(* IEC 61131-3 sources: STAR-PLC-Agent/experiments/E3/campaign_2026-11-14T074447614126+0000/PUB003/run_2026-11-14T075406993896+0000/compile_00, 1 file *)

(* ---- FB_Task.st ---- *)
FUNCTION_BLOCK FB_Task
VAR_INPUT
    Value : REAL;
    hiLevel : REAL;
    loLevel : REAL;
    hystWindow : REAL;
END_VAR
VAR_OUTPUT
    hiAlarm : BOOL := FALSE;
    loAlarm : BOOL := FALSE;
    {attribute 'analysis' := '-27'}
    error : BOOL := FALSE;
    {attribute 'analysis' := '-27'}
    status : WORD := 0;
END_VAR
VAR
    hiAlarmState : BOOL := FALSE;
    loAlarmState : BOOL := FALSE;
    span : REAL;
    hiRelease : REAL;
    loRelease : REAL;
END_VAR

span := hiLevel - loLevel;
hiRelease := hiLevel - hystWindow;
loRelease := loLevel + hystWindow;

IF loLevel >= hiLevel THEN
    error := TRUE;
    status := 16#8001;
ELSIF hystWindow >= span THEN
    error := TRUE;
    status := 16#8002;
ELSE
    error := FALSE;
    status := 0;

    IF Value > hiLevel THEN
        hiAlarmState := TRUE;
    ELSIF Value < hiRelease THEN
        hiAlarmState := FALSE;
    END_IF;

    IF Value < loLevel THEN
        loAlarmState := TRUE;
    ELSIF Value > loRelease THEN
        loAlarmState := FALSE;
    END_IF;
END_IF;

hiAlarm := hiAlarmState;
loAlarm := loAlarmState;
END_FUNCTION_BLOCK
